Staubli VAL3: HMI_safepoint.dtx

mdesc mNomSpeed
bool bBack
bool bTeach
bool bMove
string sList
string sSelPoint
bool bActive
string sTRSF[6]
string sLastPoint
mdesc mSimulate = {blend=off}
